// TIA Portal V21 export
// export: Created 2026-11-11T00:48:24.7092715Z, ExportSetting WithDefaults, DisplayName Totally Integrated Automation Portal, DisplayVersion V21 Update 3, DisplayName STEP 7 Professional, DisplayVersion V21 Update 3, DisplayName STEP 7 Safety, DisplayVersion V21, DisplayName Tech WebApplication, DisplayVersion V21, DisplayName WinCC Basic/Comfort/Advanced, DisplayVersion V21 Update 3, DisplayName WinCC Unified, DisplayVersion V21 Update 3
FUNCTION_BLOCK "FB_Scl_sl117"   // FB205, SCL
{ S7_Optimized_Access := 'TRUE' }
VERSION : 0.1
// stored: AutoNumber true, IsIECCheckEnabled false, IsRetainMemResEnabled false, MemoryReserve 100, SetENOAutomatically false, UDAEnableTagReadback false
   VAR_INPUT
      v_in : Real;
      v_sample_t : Int;
   END_VAR
   VAR_OUTPUT
      v_out : Real;
      v_err_code : Word;
   END_VAR
   VAR
      inst { S7_SetPoint := 'True'} : LEAD_LAG;
   END_VAR
BEGIN
   #inst(IN := #v_in, SAMPLE_T := #v_sample_t, OUT => #v_out, ERR_CODE => #v_err_code);
END_FUNCTION_BLOCK
